(* IEC 61131-3 sources: JingjiangMoonbox/Application/Application/任务列表/LogTask/文件存储, 4 files *)

(* ---- KS_FixedWidthStr.st ---- *)
(*@CES
Name=KS_FixedWidthStr
Type=FunctionBlock
TypeGuid=6f9dac99-8de1-4efc-8465-68ac443b7d08
Guid=54bcfd76-1fab-4aff-97a7-749ae0439a1a
HasDeclaration=True
HasImplementation=True
*)
{DECLARATION}
FUNCTION KS_FixedWidthStr : STRING
VAR_INPUT
	i_sInput: STRING;(* 输入的信息 *)
	i_iNeedWidth: INT;(* 需要的宽度 *)
END_VAR
VAR
	i: INT;
	iLen: INT;
	sResult: STRING;
END_VAR

{IMPLEMENTATION}
iLen:= LEN(i_sInput);
IF iLen>=i_iNeedWidth THEN
	sResult:= RIGHT(i_sInput, i_iNeedWidth);
ELSE
	sResult:= '';
	FOR i:=1 TO (i_iNeedWidth-iLen) BY 1 DO
		sResult:= CONCAT(sResult, '0');
	END_FOR
	sResult:= CONCAT(sResult, i_sInput);
END_IF
KS_FixedWidthStr:= sResult;

(* ---- KS_GenTimeString.st ---- *)
(*@CES
Name=KS_GenTimeString
Type=FunctionBlock
TypeGuid=6f9dac99-8de1-4efc-8465-68ac443b7d08
Guid=deb9626e-0703-4969-b954-92f6cc3bdf0c
HasDeclaration=True
HasImplementation=True
*)
{DECLARATION}
FUNCTION KS_GenTimeString : STRING
(* 输出格式yyyymmddHHMMSS[uuu]
输出yyyymmdd的dword/最大到99991231/(dword范围0~4294967295)
输出HHMMSS[uuu]的dword/最大到235959999
description:
当i_pdwDATA和i_pdwTIME都输入0时/则返回可阅读方式的字符串格式[YYYY-mm-dd HH:MM:SS.mmm]
returns:
如果SysTimeRtc.library接口调用失败会有两个特别的时间返回/以标识错误类别/分别是:'1999-12-31 23:59:59.999'和'2999-01-01 00:00:00.999';
*)
VAR_INPUT
	i_pdwDATE: POINTER TO DWORD;(* 返回日期YYYYmmdd的dword形式 *)
	i_pdwTIME: POINTER TO DWORD;(* 返回HHMMSSmmm的dword形式 *)
	i_piErrCode: POINTER TO INT;(* 错误代码/-1.SysTimeRtcHighResGet() failed/-2.SysTimeRtcConvertHighResToLocal() failed/-3. string length not equal 17 *)
END_VAR
VAR
	sResult: STRING := '';
	udiRtn: RTS_IEC_RESULT;
	stSYSTIME: SYSTIME;
	stRTS_SYSTIMEDATE: RTS_SYSTIMEDATE;
END_VAR
{IMPLEMENTATION}
IF SysTimeRtcHighResGet(stSYSTIME)=0 THEN(* 获得当前高精度UTC时间戳 *)
	IF SysTimeRtcConvertHighResToLocal(stSYSTIME, stRTS_SYSTIMEDATE)=0 THEN
		IF i_pdwDATE<>0 OR i_pdwTIME<>0 THEN(* 需要拿到日期和时间的dword类型 *)
			sResult:= CONCAT(sResult, KS_FixedWidthStr(WORD_TO_STRING(stRTS_SYSTIMEDATE.wYear), 4));
			sResult:= CONCAT(sResult, KS_FixedWidthStr(WORD_TO_STRING(stRTS_SYSTIMEDATE.wMonth), 2));
			sResult:= CONCAT(sResult, KS_FixedWidthStr(WORD_TO_STRING(stRTS_SYSTIMEDATE.wDay), 2));
			sResult:= CONCAT(sResult, KS_FixedWidthStr(WORD_TO_STRING(stRTS_SYSTIMEDATE.wHour), 2));
			sResult:= CONCAT(sResult, KS_FixedWidthStr(WORD_TO_STRING(stRTS_SYSTIMEDATE.wMinute), 2));
			sResult:= CONCAT(sResult, KS_FixedWidthStr(WORD_TO_STRING(stRTS_SYSTIMEDATE.wSecond), 2));
			sResult:= CONCAT(sResult, KS_FixedWidthStr(WORD_TO_STRING(stRTS_SYSTIMEDATE.wMilliseconds), 3));
			IF LEN(sResult)<>17 THEN(* 长度不满足要求 *)
				IF i_piErrCode<>0 THEN i_piErrCode^:= -3; END_IF
			ELSE(* 获取date和time的dword类型值 *)
				IF i_pdwDATE<>0 THEN i_pdwDATE^:= STRING_TO_DWORD(LEFT(sResult, 8)); END_IF
				IF i_pdwTIME<>0 THEN i_pdwTIME^:= STRING_TO_DWORD(RIGHT(sResult, 9)); END_IF
			END_IF
		ELSE(* 期望拿到可阅读的时间/YYYY-mm-dd HH:MM:SS.mmm格式 *)
			sResult:= CONCAT(sResult, KS_FixedWidthStr(WORD_TO_STRING(stRTS_SYSTIMEDATE.wYear), 4));
			sResult:= CONCAT(sResult, '-');
			sResult:= CONCAT(sResult, KS_FixedWidthStr(WORD_TO_STRING(stRTS_SYSTIMEDATE.wMonth), 2));
			sResult:= CONCAT(sResult, '-');
			sResult:= CONCAT(sResult, KS_FixedWidthStr(WORD_TO_STRING(stRTS_SYSTIMEDATE.wDay), 2));
			sResult:= CONCAT(sResult, ' ');
			sResult:= CONCAT(sResult, KS_FixedWidthStr(WORD_TO_STRING(stRTS_SYSTIMEDATE.wHour), 2));
			sResult:= CONCAT(sResult, ':');
			sResult:= CONCAT(sResult, KS_FixedWidthStr(WORD_TO_STRING(stRTS_SYSTIMEDATE.wMinute), 2));
			sResult:= CONCAT(sResult, ':');
			sResult:= CONCAT(sResult, KS_FixedWidthStr(WORD_TO_STRING(stRTS_SYSTIMEDATE.wSecond), 2));
			sResult:= CONCAT(sResult, '.');
			sResult:= CONCAT(sResult, KS_FixedWidthStr(WORD_TO_STRING(stRTS_SYSTIMEDATE.wMilliseconds), 3));
		END_IF
	ELSE(* SysTimeRtcConvertHighResToLocal() faield *)
		IF i_pdwDATE<>0 OR i_pdwTIME<>0 THEN
			sResult:= '29990101000000999';
		ELSE
			sResult:= '2999-01-01 00:00:00.999';
		END_IF
	END_IF
ELSE(* SysTimeRtcHighResGet() failed *)
	IF i_pdwDATE<>0 OR i_pdwTIME<>0 THEN
		sResult:= '19991231235959999';
	ELSE
		sResult:= '1999-12-31 23:59:59.999';
	END_IF
END_IF
KS_GenTimeString:= sResult;

(* ---- KS_GetTimeString.st ---- *)
(*@CES
Name=KS_GetTimeString
Type=FunctionBlock
TypeGuid=6f9dac99-8de1-4efc-8465-68ac443b7d08
Guid=2915fd67-d492-46c1-83ff-21d786551c5b
HasDeclaration=True
HasImplementation=True
*)
{DECLARATION}
FUNCTION KS_GetTimeString : STRING
VAR_INPUT
	i_iTimeFmtId: INT := TIMEFORMAT_NO_HYPHEN;
	i_xInclHMSU: BOOL := FALSE;(* 只有日期/不含具体时间部分 *)
	i_xInclMilliseconds: BOOL := FALSE;(* 包含毫秒部分/前提是i_xIncludeHMSU有效 *)
	i_pdwYMD: POINTER TO DWORD := 0;(* 年月日/最大99991231/保存数据项时如果需要/请传入合法的地址 *)
	i_pdwHMSU: POINTER TO DWORD := 0;(* 时分秒+毫秒/最大235959999/保存数据项时如果需要/请传入合法的地址 *)
END_VAR
VAR
	sResult: STRING;
	sYMD: STRING;
	sHMSU: STRING;
	stTimestamp: SYSTIME;
	stSysTimedate: RTS_SYSTIMEDATE;(* RTS_SYSTIMEDATE *)
	udiRtn: RTS_IEC_RESULT;
	asTimedateItem: ARRAY [1..7] OF STRING(10) := [7('')];

//	stSysTimedate_Rec: RTS_SYSTIMEDATE;(* RTS_SYSTIMEDATE *)

END_VAR
{IMPLEMENTATION}
udiRtn:= SysTimeRtcHighResGet(stTimestamp);(* 获得当前高精度UTC时间戳 *)
udiRtn:= SysTimeRtcConvertHighResToLocal(stTimestamp, stSysTimedate);
IF NOT g_xInitTime THEN
	g_xInitTime:= TRUE;
	SysMemCpy(ADR(g_stSysTimedate_Rec),ADR(stSysTimedate),SIZEOF(g_stSysTimedate_Rec));
END_IF
(* 年 *)
asTimedateItem[1]:= WORD_TO_STRING(stSysTimedate.wYear);

(* 月 *)
IF stSysTimedate.wMonth<10 THEN
	asTimedateItem[2]:= '0';
	asTimedateItem[2]:= CONCAT(asTimedateItem[2], WORD_TO_STRING(stSysTimedate.wMonth));
ELSE
	asTimedateItem[2]:= WORD_TO_STRING(stSysTimedate.wMonth);
END_IF

(* 日 *)
IF stSysTimedate.wDay<10 THEN
	asTimedateItem[3]:= '0';
	asTimedateItem[3]:= CONCAT(asTimedateItem[3], WORD_TO_STRING(stSysTimedate.wDay));
ELSE
	asTimedateItem[3]:= WORD_TO_STRING(stSysTimedate.wDay);
END_IF

(* 时 *)
IF g_stSysTimedate_Rec.wHour<>stSysTimedate.wHour THEN
	IF (WORD_TO_INT(stSysTimedate.wHour)-WORD_TO_INT(g_stSysTimedate_Rec.wHour)<>1) AND
		(WORD_TO_INT(stSysTimedate.wHour)-WORD_TO_INT(g_stSysTimedate_Rec.wHour)<>-23) THEN
		stSysTimedate.wHour:=  g_stSysTimedate_Rec.wHour;
	END_IF
END_IF
IF stSysTimedate.wHour<10 THEN
	asTimedateItem[4]:= '0';
	asTimedateItem[4]:= CONCAT(asTimedateItem[4], WORD_TO_STRING(stSysTimedate.wHour));
ELSE
	asTimedateItem[4]:= WORD_TO_STRING(stSysTimedate.wHour);
END_IF

(* 分 *)
IF stSysTimedate.wMinute<10 THEN
	asTimedateItem[5]:= '0';
	asTimedateItem[5]:= CONCAT(asTimedateItem[5], WORD_TO_STRING(stSysTimedate.wMinute));
ELSE
	asTimedateItem[5]:= WORD_TO_STRING(stSysTimedate.wMinute);
END_IF

(* 秒 *)
IF stSysTimedate.wSecond<10 THEN
	asTimedateItem[6]:= '0';
	asTimedateItem[6]:= CONCAT(asTimedateItem[6], WORD_TO_STRING(stSysTimedate.wSecond));
ELSE
	asTimedateItem[6]:= WORD_TO_STRING(stSysTimedate.wSecond);
END_IF

(* 毫秒 *)
IF stSysTimedate.wMilliseconds<10 THEN
	asTimedateItem[7]:= '00';
	asTimedateItem[7]:= CONCAT(asTimedateItem[7], WORD_TO_STRING(stSysTimedate.wMilliseconds));
ELSIF stSysTimedate.wMilliseconds<100 THEN
	asTimedateItem[7]:= '0';
	asTimedateItem[7]:= CONCAT(asTimedateItem[7], WORD_TO_STRING(stSysTimedate.wMilliseconds));
ELSE
	asTimedateItem[7]:= WORD_TO_STRING(stSysTimedate.wMilliseconds);
END_IF

IF i_iTimeFmtId=TIMEFORMAT_NO_HYPHEN THEN(* yyyymmdd[HHMMSS[uuu]] *)
	sResult:= asTimedateItem[1];
	sResult:= CONCAT(sResult, asTimedateItem[2]);
	sResult:= CONCAT(sResult, asTimedateItem[3]);
	IF i_xInclHMSU THEN
		sResult:= CONCAT(sResult, asTimedateItem[4]);
		sResult:= CONCAT(sResult, asTimedateItem[5]);
		sResult:= CONCAT(sResult, asTimedateItem[6]);
		IF i_xInclMilliseconds THEN
			sResult:= CONCAT(sResult, asTimedateItem[7]);
		END_IF
	END_IF
ELSIF i_iTimeFmtId=TIMEFORMAT_HYPHEN_COLON THEN(* yyyy-mm-dd[ HH:MM:SS[.uuu]] *)
	sResult:= asTimedateItem[1];
	sResult:= CONCAT(sResult, '-'); sResult:= CONCAT(sResult, asTimedateItem[2]);
	sResult:= CONCAT(sResult, '-'); sResult:= CONCAT(sResult, asTimedateItem[3]);
	IF i_xInclHMSU THEN
		sResult:= CONCAT(sResult, ' '); sResult:= CONCAT(sResult, asTimedateItem[4]);
		sResult:= CONCAT(sResult, ':'); sResult:= CONCAT(sResult, asTimedateItem[5]);
		sResult:= CONCAT(sResult, ':'); sResult:= CONCAT(sResult, asTimedateItem[6]);
		IF i_xInclMilliseconds THEN
			sResult:= CONCAT(sResult, '.'); sResult:= CONCAT(sResult, asTimedateItem[7]);
		END_IF
	END_IF
ELSIF i_iTimeFmtId=TIMEFORMAT_MMDD THEN(* mmdd *)
	sResult:= asTimedateItem[2];
	sResult:= CONCAT(sResult, asTimedateItem[3]);
ELSIF i_iTimeFmtId=TIMEFORMAT_MMDDHH THEN(* mmddHH *)
	sResult:= asTimedateItem[2];
	sResult:= CONCAT(sResult, asTimedateItem[3]);
	sResult:= CONCAT(sResult, asTimedateItem[4]);
ELSE(* include [i_iTimeFmtId=TIMEFORMAT_HYPHEN_DOT](* yyyy.mm.dd[.HHMMSS[_uuu]] *) *)
	sResult:= asTimedateItem[1];
	sResult:= CONCAT(sResult, '.'); sResult:= CONCAT(sResult, asTimedateItem[2]);
	sResult:= CONCAT(sResult, '.'); sResult:= CONCAT(sResult, asTimedateItem[3]);
	IF i_xInclHMSU THEN
		sResult:= CONCAT(sResult, '.'); sResult:= CONCAT(sResult, asTimedateItem[4]);
		sResult:= CONCAT(sResult, asTimedateItem[5]);
		sResult:= CONCAT(sResult, asTimedateItem[6]);
		IF i_xInclMilliseconds THEN
			sResult:= CONCAT(sResult, '_');
			sResult:= CONCAT(sResult, asTimedateItem[7]);
		END_IF
	END_IF
END_IF
IF i_pdwYMD<>0 THEN(* 年月日 *)
	sYMD:= asTimedateItem[1];
	sYMD:= CONCAT(sYMD, asTimedateItem[2]);
	sYMD:= CONCAT(sYMD, asTimedateItem[3]);
	i_pdwYMD^:= STRING_TO_DWORD(sYMD);
END_IF
IF i_pdwHMSU<>0 THEN(* 时分秒+毫秒 *)
	sHMSU:= asTimedateItem[4];
	sHMSU:= CONCAT(sHMSU, asTimedateItem[5]);
	sHMSU:= CONCAT(sHMSU, asTimedateItem[6]);
	sHMSU:= CONCAT(sHMSU, asTimedateItem[7]);
	i_pdwHMSU^:= STRING_TO_DWORD(sHMSU);
END_IF
SysMemCpy(ADR(g_stSysTimedate_Rec),ADR(stSysTimedate),SIZEOF(g_stSysTimedate_Rec));

KS_GetTimeString:= sResult;

(* ---- KS_FB_TravelFileService.st ---- *)
(*@CES
Name=KS_FB_TravelFileService
Type=FunctionBlock
TypeGuid=6f9dac99-8de1-4efc-8465-68ac443b7d08
Guid=9263010e-7967-4803-a57a-bbeff11eb4c3
HasDeclaration=True
HasImplementation=True
*)
{DECLARATION}
FUNCTION_BLOCK KS_FB_TravelFileService
(* 运行文件服务/包含日志和实时保存的数据 *)
VAR_INPUT
	i_xEn: BOOL;(* 总使能标志 *)
	i_xLog_need: BOOL;(* 置TRUE表示需要保存日志 *)
	i_xDat_need: BOOL;(* 置TRUE表示需要保存数据/可以绑定印刷条件等等 *)
	i_xReq_safeclose: BOOL;(* 请求安全关闭文件/关注本地驱动器的缺相和欠压报警标志 *)
	i_pxRst_protect: POINTER TO BOOL;(* 复位紧急保护的标志/由于在驱动器出现缺相或者欠压报警会触发紧急关闭文件/一旦出现报警/必须置复位标志才能继续保存新的文件 *)
(*deprecate@2025.8.27.164512/han.dp
	i_pstStTravelLogRec: POINTER TO StTravelLogRec;(* 完整日志区域/对应g_apstStTravelLogRec[1] *)
*)
	i_pstStTravelDataRec: POINTER TO StTravelDataRec;(* 后台记录的运行数据区域/对应g_pstStTravelDataRec *)
	i_pstStSysParam: POINTER TO StSysParam;
END_VAR
VAR_OUTPUT
	o_xEno: BOOL;
	o_sFilename_datfile: STRING;
	o_sFilename_logfile: STRING;
	o_iErNo_datfile: INT;
	o_iErNo_logfile: INT;
	o_xFileClosed_BecauseEmergency: BOOL := FALSE;
END_VAR
VAR
	sFilename: STRING;
	uiR_tmp: UINT;
	uiW_tmp: UINT;
	dwTmp: DWORD;
	dwBytesWrote_total: DWORD;
	dwHdl_logfile: DWORD := 0;(* 日志文件句柄 *)
	dwHdl_datfile: DWORD := 0;(* 数据文件句柄 *)
	xReqCloseLogfile_tmp: BOOL;
	xReqCloseDatfile_tmp: BOOL;
	iMaxDataItemsNum: INT;
	LINETAIL: BYTE := 13;(* 文本换行 *)
	pResult: RTS_IEC_RESULT;
	iRtn : INT;
	sFileName_test: STRING;
	time1:TIME;
	time2:TIME;
	adwNumByteOfFile : ARRAY[1..10] OF DWORD;
	sYMDHtemp:STRING;
	iN: INT;
	uiIdx_R_tmp:UINT;
	udiTmpOfst: UDINT;
	uiTmpRdNum: UINT;(* 2025.10.14.142248/han.dp/读取数量临时变量 *)

	pstStGrpParam_Save : POINTER TO StGrpParam_Save;

END_VAR
VAR CONSTANT
	DATFILE_MAXBYTES: DWORD := 16777216;(* 16*1024*1024字节/16MB *)
	//DATFILE_MAXBYTES: DWORD := 33554432;(* 32*1024*1024字节/16MB *)
END_VAR
{IMPLEMENTATION}
o_xEno:= i_xEn;
o_iErNo_datfile:= 0;
o_iErNo_logfile:= 0;
xReqCloseLogfile_tmp:= FALSE;
xReqCloseDatfile_tmp:= FALSE;
IF i_xEn THEN
	pstStGrpParam_Save := ADR(i_pstStSysParam^.astStGrpParam_Save[1]);
	(* 一旦紧急情况发生/开始触发文件安全关闭 *)
	IF i_xReq_safeclose AND (NOT o_xFileClosed_BecauseEmergency) THEN
		o_xFileClosed_BecauseEmergency:= TRUE;

	END_IF
	IF o_xFileClosed_BecauseEmergency THEN
		xReqCloseLogfile_tmp:= TRUE;
		xReqCloseDatfile_tmp:= TRUE;
	END_IF

	(* 可以人工启动文件保存功能 *)
	IF i_pxRst_protect<>0 THEN
		IF i_pxRst_protect^ AND (NOT i_xReq_safeclose) AND o_xFileClosed_BecauseEmergency THEN
			o_xFileClosed_BecauseEmergency:= FALSE;
		END_IF
		i_pxRst_protect^:= FALSE;(* 2023.7.26.175651/han.dp *)
	END_IF

	(* 所有的文件操作都需要在非紧急情况下进行/紧急情况一般为缺相或者欠压等供电异常状态/防止对DOM盘和OS文件造成破坏 *)
	IF NOT o_xFileClosed_BecauseEmergency THEN

(* deprecated@2025.8.27.161857/han.dp
		(* -------------------------------------------------- *)
		(* 处理日志 *)
		(* -------------------------------------------------- *)
		IF i_xLog_need THEN(* 需要保存日志 *)
			IF i_pstStTravelLogRec<>0 AND dwHdl_logfile<>0 THEN(* 写数据 *)
				uiR_tmp:= i_pstStTravelLogRec^.uiIndex_Rd;(* 读取位置 *)
				uiW_tmp:= i_pstStTravelLogRec^.uiIndex_Wr;(* 写入位置 *)
				iMaxDataItemsNum:= DWORD_TO_INT(SIZEOF(i_pstStTravelLogRec^.astStTravelLogItem)/SIZEOF(i_pstStTravelLogRec^.astStTravelLogItem[1]));(* 位置上限 *)
				IF (uiR_tmp>=1 AND uiR_tmp<=iMaxDataItemsNum) AND (uiW_tmp>=1 AND uiW_tmp<=iMaxDataItemsNum) THEN
					WHILE uiR_tmp<>uiW_tmp DO
						adwNumByteOfFile[1] := SysFileWrite(dwHdl_logfile,
							ADR(i_pstStTravelLogRec^.astStTravelLogItem[uiR_tmp].sInfo),
							LEN(i_pstStTravelLogRec^.astStTravelLogItem[uiR_tmp].sInfo), 0);
						adwNumByteOfFile[2] := SysFileWrite(dwHdl_logfile, ADR(LINETAIL), SIZEOF(LINETAIL), 0);

						uiR_tmp:= uiR_tmp+1;
						IF uiR_tmp>iMaxDataItemsNum THEN uiR_tmp:= uiR_tmp-iMaxDataItemsNum; END_IF

							uiIdx_R_tmp:= uiR_tmp;
							FOR iN:=1 TO MIN(MAX_LOG_ITEM_VIEW,GC_LOG_ITEM_MAX_NUM) BY 1 DO
								uiIdx_R_tmp:= uiIdx_R_tmp-1;
								IF uiIdx_R_tmp<1 THEN
									uiIdx_R_tmp:= uiIdx_R_tmp+GC_LOG_ITEM_MAX_NUM;
									IF NOT gvl.g_pstStTravelLogRec^.xOverwrite THEN(* 未过圈/不要复制之前的 *)
										EXIT;
									END_IF
								END_IF
								gvl.g_astStTravelLogItem_view[iN]:= gvl.g_pstStTravelLogRec^.astStTravelLogItem[uiIdx_R_tmp];
							END_FOR
						END_WHILE

					i_pstStTravelLogRec^.uiIndex_Rd:= uiR_tmp;
				ELSE
					i_pstStTravelLogRec^.uiIndex_Rd:= 1;
					i_pstStTravelLogRec^.uiIndex_Wr:= 1;
				END_IF
			ELSIF i_pstStTravelLogRec<>0 THEN(* 创建文件 *)
				sFilename:= PATH_HOME_LOG;
				sFilename:= CONCAT(sFilename, KS_GetTimeString(TIMEFORMAT_NO_HYPHEN,FALSE,FALSE,0,0));
				sFilename:= CONCAT(sFilename, '.txt');
				dwHdl_logfile:= SysFileOpen(sFilename, SysFile.AM_APPEND_PLUS, ADR(pResult));(* 以追加方式打开文件(未使用AM_WRITE模式)/失败了就会创建新的文件 *)
				IF dwHdl_logfile<>0 THEN o_sFilename_logfile:= sFilename; END_IF
			ELSE(* 关闭文件 *)
				o_iErNo_logfile:= -1;
				xReqCloseLogfile_tmp:= TRUE;
			END_IF
		ELSE xReqCloseLogfile_tmp:= TRUE; END_IF
*)

		(* -------------------------------------------------- *)
		(* 处理数据 *)
		(* -------------------------------------------------- *)
		IF i_xDat_need THEN(* 需要保存数据 *)
			IF i_pstStTravelDataRec<>0 AND dwHdl_datfile<>0 THEN(* 写数据 *)
				uiR_tmp:= i_pstStTravelDataRec^.uiRD;
				uiW_tmp:= i_pstStTravelDataRec^.uiWR;
				iMaxDataItemsNum:= DWORD_TO_INT(SIZEOF(i_pstStTravelDataRec^.astStTravelDataItem)/SIZEOF(i_pstStTravelDataRec^.astStTravelDataItem[1]));
				IF (uiR_tmp>=1 AND uiR_tmp<=iMaxDataItemsNum) AND (uiW_tmp>=1 AND uiW_tmp<=iMaxDataItemsNum) THEN
					WHILE uiR_tmp<>uiW_tmp DO

(* 2025.10.14.142930/han.dp/
/ 在写文件前把这个fifo给网络上也写一份
/ udp自动会搬到金刚主机
/ 原先的存储逻辑就会触发生效
/ 以FE_yyyymmdd.MIX文件呈现
*)
udiTmpOfst:= 0;
uiTmpRdNum:= i_pstStTravelDataRec^.astStTravelDataItem[uiR_tmp].uiValidBytesNum;
WHILE uiTmpRdNum>=1020 DO
	KS_PushDataToFifo(TRUE,
		ADR(i_pstStTravelDataRec^.astStTravelDataItem[uiR_tmp].abyPayload)+udiTmpOfst,
		1020,
		g_pstStUdpOnlySendFifo);
	uiTmpRdNum:= uiTmpRdNum-1020;
	udiTmpOfst:= udiTmpOfst+1020;
END_WHILE
IF uiTmpRdNum<>0 THEN
	KS_PushDataToFifo(TRUE,
		ADR(i_pstStTravelDataRec^.astStTravelDataItem[uiR_tmp].abyPayload)+udiTmpOfst,
		uiTmpRdNum,
		g_pstStUdpOnlySendFifo);
END_IF

						IF pstStGrpParam_Save^.dwExtBitCtlFlag.22 THEN
							dwTmp:= SysFileWrite(dwHdl_datfile,
								ADR(i_pstStTravelDataRec^.astStTravelDataItem[uiR_tmp].abyPayload),
								i_pstStTravelDataRec^.astStTravelDataItem[uiR_tmp].uiValidBytesNum, ADR(pResult));
						END_IF
						uiR_tmp:= uiR_tmp+1;
						IF uiR_tmp>iMaxDataItemsNum THEN uiR_tmp:= uiR_tmp-iMaxDataItemsNum; END_IF
						dwBytesWrote_total:= dwBytesWrote_total+dwTmp;
						IF dwBytesWrote_total>=DATFILE_MAXBYTES THEN(* 文件写够约定的大小就切换/请注意:要保证最后1包数据是完整的/并不是按照文件严格的定长来切换文件的 *)
							xReqCloseDatfile_tmp:= TRUE;
							EXIT;
						END_IF
					END_WHILE
					i_pstStTravelDataRec^.uiRD:= uiR_tmp;
				ELSE
					i_pstStTravelDataRec^.uiRD:= 1;
					i_pstStTravelDataRec^.uiWR:= 1;
				END_IF
			ELSIF i_pstStTravelDataRec<>0 THEN(* 创建文件 *)
				(*sYMDHtemp:=KS_GetTimeString(TIMEFORMAT_MMDDHH, FALSE, FALSE);
				PATH_HOME_DATA:=concat('/opt/codesyscontrol/kesai/data/',KS_GetTimeString(TIMEFORMAT_MMDDHH,TRUE,FALSE,0,0));
				PATH_HOME_DATA:=concat(PATH_HOME_DATA,'/');
				*)
				sFilename:= PATH_HOME_DATA;
				sFilename:= CONCAT(sFilename, KS_GetTimeString(TIMEFORMAT_NO_HYPHEN,TRUE,FALSE,0,0));(* 精确到s就可以 *)

				//使用新系统之后路径发生变化  /opt/codesyscontrol/---->/data/
				//sFilename:= MID(sFilename,41,1);
				sFilename:= MID(sFilename,27,1);
				sFilename:= CONCAT(sFilename,'/');
				sFilename:= CONCAT(sFilename, KS_GetTimeString(TIMEFORMAT_NO_HYPHEN,TRUE,FALSE,0,0));(* 精确到s就可以 *)

				sFilename:= CONCAT(sFilename, '.MIX');
				dwBytesWrote_total:= 0;(* 总计写入字节数量清零 *)
				dwHdl_datfile:= SysFileOpen(sFilename, SysFile.AM_WRITE, ADR(pResult));
				IF dwHdl_datfile<>0 THEN o_sFilename_datfile:= sFilename; END_IF
			ELSE(* 关闭文件 *)
				o_iErNo_datfile:= -1;
				xReqCloseDatfile_tmp:= TRUE;
			END_IF
		ELSE xReqCloseDatfile_tmp:= TRUE; END_IF
	END_IF

ELSE
	xReqCloseLogfile_tmp:= TRUE;
	xReqCloseDatfile_tmp:= TRUE;
END_IF

IF xReqCloseLogfile_tmp AND dwHdl_logfile<>0 THEN(* 关闭日志文件 *)
	SysFileClose(dwHdl_logfile);
	dwHdl_logfile:= 0;
	o_sFilename_logfile:= '';
END_IF

IF xReqCloseDatfile_tmp AND dwHdl_datfile<>0 THEN(* 关闭数据文件 *)
	SysFileClose(dwHdl_datfile);
	dwHdl_datfile:= 0;
	o_sFilename_datfile:= '';
END_IF
